KUKA KRL data list: folge11.dat

&ACCESS RVP
&REL 1
&COMMENT bt2krl sim data Folge 11 plan 16#4F80
DEFDAT FOLGE11
   ; Generated by bt2krl 0.1.0 from bt2plc plan bt_1792076124_welding_cell_2_small (cell welding_cell_2_small), PLAN_ID 16#4F80
   ; Robot robot1 (R1), controller robot1, model KR240R2900_ULTRA, joint mapping identity
   ; Profile sim (bt2plc simulator telegram). NEVER install on a VW KS24 robot:
   ; its signals collide with the VW standard (Fertigmeldung, interlocks, PRG_NR).
   ; Do not edit: regenerate with bt2krl (plain KRL, no inline forms).
   EXT BAS (BAS_COMMAND :IN,REAL :IN )
   DECL INT PLAN_ID=20352
   DECL AXIS P1={A1 0.0,A2 -90.0,A3 90.0,A4 0.0,A5 0.0,A6 0.0}
   DECL AXIS P2={A1 -0.5763,A2 -90.0384,A3 90.0828,A4 -0.2659,A5 0.4589,A6 0.5219}
   DECL AXIS P3={A1 -3.6018,A2 -90.2401,A3 90.5176,A4 -1.662,A5 2.8686,A6 3.2621}
   DECL AXIS P4={A1 -7.0597,A2 -90.4706,A3 91.0145,A4 -3.2576,A5 5.6225,A6 6.3939}
   DECL AXIS P5={A1 -14.4077,A2 -90.9605,A3 92.0704,A4 -6.6481,A5 11.4747,A6 13.0489}
   DECL AXIS P6={A1 -20.7472,A2 -91.3831,A3 92.9814,A4 -9.5733,A5 16.5236,A6 18.7906}
   DECL AXIS P7={A1 -32.4177,A2 -92.1611,A3 94.6584,A4 -14.9583,A5 25.8182,A6 29.3603}
   DECL AXIS P8={A1 -41.6387,A2 -92.7758,A3 95.9835,A4 -19.2132,A5 33.1622,A6 37.7118}
   DECL AXIS P9={A1 -61.738,A2 -94.1157,A3 98.8717,A4 -28.4875,A5 49.1697,A6 55.9155}
   DECL AXIS P10={A1 -74.2731,A2 -94.9514,A3 100.673,A4 -34.2715,A5 59.153,A6 67.2684}
   DECL AXIS P11={A1 -81.1891,A2 -95.4124,A3 101.6668,A4 -37.4627,A5 64.661,A6 73.5321}
   DECL AXIS P12={A1 -86.9524,A2 -95.7966,A3 102.495,A4 -40.122,A5 69.2511,A6 78.7518}
   DECL AXIS P13={A1 -93.4361,A2 -96.2288,A3 103.4267,A4 -43.1138,A5 74.4149,A6 84.6241}
   DECL AXIS P14={A1 -96.3178,A2 -96.4209,A3 103.8409,A4 -44.4434,A5 76.7099,A6 87.234}
   DECL AXIS P15={A1 -98.4791,A2 -96.565,A3 104.1514,A4 -45.4407,A5 78.4313,A6 89.1915}
   DECL AXIS P16={A1 -98.6233,A2 -95.6972,A3 108.0019,A4 -46.2938,A5 75.2694,A6 92.7921}
   DECL AXIS P17={A1 -98.6233,A2 -95.6972,A3 108.0016,A4 -46.2937,A5 75.2695,A6 92.7919}
   DECL AXIS P18={A1 -98.768,A2 -96.5112,A3 104.0441,A4 -45.2543,A5 78.6321,A6 89.1332}
   DECL AXIS P19={A1 -99.9229,A2 -96.0049,A3 103.022,A4 -43.2364,A5 79.319,A6 87.626}
   DECL AXIS P20={A1 -102.232,A2 -94.9926,A3 100.9784,A4 -39.2015,A5 80.6922,A6 84.6124}
   DECL AXIS P21={A1 -105.6955,A2 -93.4743,A3 97.9132,A4 -33.1497,A5 82.752,A6 80.0923}
   DECL AXIS P22={A1 -115.4301,A2 -89.2068,A3 89.2978,A4 -16.1398,A5 88.5412,A6 67.3878}
   DECL AXIS P23={A1 -119.4707,A2 -87.4355,A3 85.7218,A4 -9.0795,A5 90.9442,A6 62.1145}
   DECL AXIS P24={A1 -122.357,A2 -86.1702,A3 83.1674,A4 -4.0361,A5 92.6607,A6 58.3477}
   DECL AXIS P25={A1 -124.089,A2 -85.4109,A3 81.6346,A4 -1.0097,A5 93.6908,A6 56.0873}
   DECL AXIS P26={A1 -124.6667,A2 -85.1576,A3 81.1233,A4 -0.0002,A5 94.0343,A6 55.3333}
   DECL AXIS P27={A1 -124.6668,A2 -85.1195,A3 85.5727,A4 0.0,A5 89.5468,A6 55.3331}
   DECL AXIS P28={A1 -124.6668,A2 -85.1195,A3 85.5727,A4 0.0,A5 89.5468,A6 55.3331}
   DECL AXIS P29={A1 -124.5299,A2 -85.1588,A3 81.1836,A4 -0.2276,A5 93.9611,A6 55.5086}
   DECL AXIS P30={A1 -123.4341,A2 -85.1682,A3 81.6672,A4 -2.0488,A5 93.3737,A6 56.9128}
   DECL AXIS P31={A1 -119.7353,A2 -85.2001,A3 83.2994,A4 -8.1962,A5 91.3914,A6 61.6524}
   DECL AXIS P32={A1 -115.8994,A2 -85.2332,A3 84.9922,A4 -14.5715,A5 89.3355,A6 66.5678}
   DECL AXIS P33={A1 -108.3645,A2 -85.2981,A3 88.3174,A4 -27.0948,A5 85.2971,A6 76.2232}
   DECL AXIS P34={A1 -103.9802,A2 -85.3359,A3 90.2522,A4 -34.3816,A5 82.9473,A6 81.8413}
   DECL AXIS P35={A1 -100.6918,A2 -85.3643,A3 91.7033,A4 -39.8468,A5 81.185,A6 86.0551}
   DECL AXIS P36={A1 -98.4995,A2 -85.3832,A3 92.6708,A4 -43.4904,A5 80.01,A6 88.8643}
   DECL AXIS P37={A1 -97.2662,A2 -85.3938,A3 93.2151,A4 -45.5403,A5 79.349,A6 90.4447}
   DECL AXIS P38={A1 -97.2661,A2 -84.546,A3 96.8787,A4 -46.2424,A5 76.208,A6 93.7588}
   DECL AXIS P39={A1 -97.2661,A2 -84.5461,A3 96.8785,A4 -46.2423,A5 76.2082,A6 93.7586}
   DECL AXIS P40={A1 -97.2662,A2 -85.3937,A3 93.215,A4 -45.5401,A5 79.3491,A6 90.4448}
   DECL AXIS P41={A1 -98.5436,A2 -84.7944,A3 92.4187,A4 -43.2914,A5 80.4888,A6 90.3788}
   DECL AXIS P42={A1 -102.3741,A2 -82.997,A3 90.0306,A4 -36.5482,A5 83.9065,A6 90.1807}
   DECL AXIS P43={A1 -106.3461,A2 -81.1333,A3 87.5543,A4 -29.5559,A5 87.4504,A6 89.9755}
   DECL AXIS P44={A1 -114.4316,A2 -77.3393,A3 82.5135,A4 -15.3219,A5 94.6647,A6 89.5575}
   DECL AXIS P45={A1 -127.4092,A2 -71.2499,A3 74.4228,A4 7.5239,A5 106.2437,A6 88.8868}
   DECL AXIS P46={A1 -134.642,A2 -67.8561,A3 69.9136,A4 20.2566,A5 112.6971,A6 88.5129}
   DECL AXIS P47={A1 -139.3218,A2 -65.6602,A3 66.9961,A4 28.495,A5 116.8726,A6 88.2711}
   DECL AXIS P48={A1 -141.0233,A2 -64.8619,A3 65.9353,A4 31.4903,A5 118.3907,A6 88.1831}
   DECL AXIS P49={A1 -141.5902,A2 -64.5958,A3 65.5821,A4 32.4882,A5 118.8964,A6 88.1537}
   DECL AXIS P50={A1 -141.5902,A2 -64.1977,A3 69.4969,A4 31.3229,A5 115.2344,A6 85.5943}
   DECL AXIS P51={A1 -141.5902,A2 -64.1977,A3 69.4969,A4 31.3229,A5 115.2344,A6 85.5943}
   DECL AXIS P52={A1 -141.5902,A2 -64.5958,A3 65.5819,A4 32.4883,A5 118.8965,A6 88.1538}
   DECL AXIS P53={A1 -141.5902,A2 -64.5958,A3 65.5819,A4 32.4883,A5 118.8965,A6 88.1538}
   DECL AXIS P54={A1 -141.5389,A2 -64.5129,A3 65.4513,A4 32.5266,A5 118.9019,A6 88.0807}
   DECL AXIS P55={A1 -141.1278,A2 -63.8492,A3 64.4058,A4 32.8332,A5 118.9443,A6 87.4952}
   DECL AXIS P56={A1 -140.3054,A2 -62.5213,A3 62.3142,A4 33.4466,A5 119.0293,A6 86.3241}
   DECL AXIS P57={A1 -137.3748,A2 -57.7897,A3 54.8613,A4 35.6324,A5 119.3322,A6 82.1507}
   DECL AXIS P58={A1 -136.7576,A2 -56.7933,A3 53.2917,A4 36.0928,A5 119.396,A6 81.2719}
   DECL AXIS P59={A1 -136.5518,A2 -56.4609,A3 52.7682,A4 36.2463,A5 119.4173,A6 80.9787}
   DECL AXIS P60={A1 -136.5518,A2 -56.3896,A3 57.1431,A4 34.8931,A5 115.7998,A6 78.0604}
   DECL AXIS P61={A1 -136.5518,A2 -56.3896,A3 57.1433,A4 34.893,A5 115.7996,A6 78.0602}
   DECL AXIS P62={A1 -136.5518,A2 -56.4608,A3 52.7683,A4 36.2463,A5 119.4171,A6 80.9785}
   DECL AXIS P63={A1 -136.4239,A2 -56.609,A3 52.8988,A4 35.9634,A5 119.2338,A6 80.8135}
   DECL AXIS P64={A1 -136.0395,A2 -57.0546,A3 53.2923,A4 35.1125,A5 118.6821,A6 80.3169}
   DECL AXIS P65={A1 -134.5043,A2 -58.8339,A3 54.8633,A4 31.7146,A5 116.4789,A6 78.3338}
   DECL AXIS P66={A1 -131.9461,A2 -61.7991,A3 57.4812,A4 26.0523,A5 112.8075,A6 75.0291}
   DECL AXIS P67={A1 -126.4462,A2 -68.1738,A3 63.1095,A4 13.8788,A5 104.9143,A6 67.9243}
   DECL AXIS P68={A1 -123.3733,A2 -71.7354,A3 66.254,A4 7.0774,A5 100.5043,A6 63.9548}
   DECL AXIS P69={A1 -121.327,A2 -74.1072,A3 68.3481,A4 2.5481,A5 97.5676,A6 61.3114}
   DECL AXIS P70={A1 -120.3038,A2 -75.2932,A3 69.3952,A4 0.2833,A5 96.0991,A6 59.9895}
   DECL AXIS P71={A1 -120.1758,A2 -75.5343,A3 74.1378,A4 0.0,A5 91.3965,A6 59.8242}
   DECL AXIS P72={A1 -120.1758,A2 -75.5343,A3 74.138,A4 0.0,A5 91.3963,A6 59.8242}
   DECL AXIS P73={A1 -120.0501,A2 -75.0529,A3 68.9841,A4 0.0,A5 96.0689,A6 59.9499}
   DECL AXIS P74={A1 -119.3897,A2 -73.0116,A3 66.1364,A4 0.0,A5 96.8751,A6 60.6103}
   DECL AXIS P75={A1 -117.77,A2 -68.0044,A3 59.1515,A4 0.0,A5 98.8529,A6 62.23}
   DECL AXIS P76={A1 -117.1408,A2 -66.0594,A3 56.4382,A4 0.0,A5 99.6212,A6 62.8592}
   DECL AXIS P77={A1 -116.6688,A2 -64.6003,A3 54.4028,A4 0.0,A5 100.1975,A6 63.3312}
   DECL AXIS P78={A1 -116.6372,A2 -64.9407,A3 59.4329,A4 0.0,A5 95.5078,A6 63.3628}
   DECL AXIS P79={A1 -116.6372,A2 -64.9407,A3 59.4329,A4 0.0,A5 95.5078,A6 63.3628}
   DECL AXIS P80={A1 -116.6372,A2 -64.5028,A3 54.267,A4 0.0,A5 100.2358,A6 63.3628}
   DECL AXIS P81={A1 -115.3155,A2 -64.7917,A3 54.6716,A4 0.0,A5 99.1002,A6 62.6447}
   DECL AXIS P82={A1 -112.9672,A2 -65.305,A3 55.3911,A4 0.0,A5 97.0821,A6 61.3691}
   DECL AXIS P83={A1 -109.445,A2 -66.075,A3 56.4701,A4 0.0,A5 94.0551,A6 59.4556}
   DECL AXIS P84={A1 -101.9608,A2 -67.7111,A3 58.7631,A4 0.0,A5 87.6233,A6 55.3898}
   DECL AXIS P85={A1 -95.5039,A2 -69.1226,A3 60.7412,A4 0.0,A5 82.0744,A6 51.8821}
   DECL AXIS P86={A1 -87.8731,A2 -70.7907,A3 63.079,A4 0.0,A5 75.5166,A6 47.7368}
   DECL AXIS P87={A1 -74.226,A2 -73.774,A3 67.26,A4 0.0,A5 63.7885,A6 40.323}
   DECL AXIS P88={A1 -42.4196,A2 -80.7269,A3 77.0042,A4 0.0,A5 36.4547,A6 23.0443}
   DECL AXIS P89={A1 -33.0183,A2 -82.7821,A3 79.8844,A4 0.0,A5 28.3754,A6 17.9371}
   DECL AXIS P90={A1 -24.8008,A2 -84.5785,A3 82.4019,A4 0.0,A5 21.3134,A6 13.473}
   DECL AXIS P91={A1 -17.7572,A2 -86.1182,A3 84.5599,A4 0.0,A5 15.2602,A6 9.6465}
   DECL AXIS P92={A1 -9.3927,A2 -87.9467,A3 87.1224,A4 0.0,A5 8.0719,A6 5.1026}
   DECL AXIS P93={A1 -5.2838,A2 -88.845,A3 88.3813,A4 0.0,A5 4.5407,A6 2.8704}
   DECL AXIS P94={A1 -2.3487,A2 -89.4866,A3 89.2805,A4 0.0,A5 2.0184,A6 1.2759}
   DECL AXIS P95={A1 -0.5875,A2 -89.8716,A3 89.82,A4 0.0,A5 0.5049,A6 0.3191}
   DECL AXIS P96={A1 -0.0001,A2 -90.0,A3 90.0,A4 0.0,A5 0.0001,A6 0.0001}
   DECL AXIS P97={A1 0.0,A2 -90.0,A3 90.0,A4 0.0,A5 0.0,A6 0.0}
   DECL AXIS P98={A1 0.0,A2 -90.0,A3 90.0,A4 0.0,A5 0.0,A6 0.0}
   DECL AXIS P99={A1 0.0,A2 -90.0,A3 90.0,A4 0.0,A5 0.0,A6 0.0}
ENDDAT
